(* IEC 61131-3 sources: sis-interlock-demo/src/GVLs/Generated, 3 files *)

(* ---- GVL_Sis.gvl.st ---- *)
// AUTO-GENERATED by cemgen 1.0.0 — не редактировать: правьте матрицу и запустите
//   python -m cemgen generate <файл матрицы .csv или .xlsx>
// Матрица: SIS-V101-CEM, объект V-101, ревизия B от 2026-10-19, SHA-256 сетки df2ed4841a9453ca
// Назначение: экземпляры ПАЗ объекта V-101: источник времени, журнал событий, приложение ПАЗ и
//             команды HMI (ST_SisCmd). Вызов — PRG_Sis.
// Автор:      kr0nsch; код — генератор cemgen
// Версия:     1.0.0
// Документ:   docs/DESIGN.md, раздел «10. Генератор cemgen»; docs/cause_effect_matrix.md
// ВНИМАНИЕ:   код демонстрационный и не предназначен для систем безопасности. Реальная ПАЗ требует
//             определения SIL, сертифицированных аппаратных и программных средств и валидации по
//             ГОСТ Р МЭК 61511.
{attribute 'qualified_only'}
VAR_GLOBAL
    fbTime : PL.FB_SystemTime;   // монотонное время LTIME (PL.I_TimeSource)
    fbLog  : FB_SisEventLog;     // журнал событий ПАЗ, кольцо GVL_Const.SIS_LOG_SIZE
    fbApp  : FB_SisApp;          // ПАЗ объекта: привязка, голосование, матрица, выходы
    stCmd  : ST_SisCmd;          // команды HMI: сброс, пусковые обходы, байпасы каналов
END_VAR

(* ---- GVL_SisCfg.gvl.st ---- *)
// AUTO-GENERATED by cemgen 1.0.0 — не редактировать: правьте матрицу и запустите
//   python -m cemgen generate <файл матрицы .csv или .xlsx>
// Матрица: SIS-V101-CEM, объект V-101, ревизия B от 2026-10-19, SHA-256 сетки df2ed4841a9453ca
// Назначение: конфигурация ПАЗ объекта V-101 из матрицы причин и следствий: номера причин и
//             следствий, шкалы датчиков, матрица CEM_CFG (с CRC) и группы голосования VOTE_CFG.
//             VAR_GLOBAL CONSTANT: с HMI не меняется (решение D-09), правка — только через матрицу
//             и генератор.
// Автор:      kr0nsch; код — генератор cemgen
// Версия:     1.0.0
// Документ:   docs/DESIGN.md, раздел «10. Генератор cemgen»; docs/cause_effect_matrix.md
// ВНИМАНИЕ:   код демонстрационный и не предназначен для систем безопасности. Реальная ПАЗ требует
//             определения SIL, сертифицированных аппаратных и программных средств и валидации по
//             ГОСТ Р МЭК 61511.
{attribute 'qualified_only'}
VAR_GLOBAL CONSTANT
    // Номера причин: индекс i строки матрицы, бит маски i − 1
    CAUSE_PSHH101       : UINT := 1;   // Давление в V-101 аварийно высокое
    CAUSE_PSLL101       : UINT := 2;   // Давление в V-101 аварийно низкое
    CAUSE_LSHH102       : UINT := 3;   // Уровень жидкости в V-101 аварийно высокий
    CAUSE_LSLL102       : UINT := 4;   // Уровень жидкости в V-101 аварийно низкий
    CAUSE_TSHH103       : UINT := 5;   // Температура жидкости в V-101 аварийно высокая
    CAUSE_ASHH104       : UINT := 6;   // Загазованность у V-101 аварийно высокая
    CAUSE_BSH105        : UINT := 7;   // Пожар у V-101
    CAUSE_HS106         : UINT := 8;   // Аварийный останов кнопкой
    CAUSE_PSLL108       : UINT := 9;   // Давление воздуха КИП аварийно низкое
    CAUSE_ESL109        : UINT := 10;   // Потеря напряжения щита 0,4 кВ
    CAUSE_COUNT         : UINT := 10;   // причин в матрице
    // Номера следствий: индекс j столбца матрицы
    EFFECT_ESDV101      : UINT := 1;   // Клапан-отсекатель на входе V-101
    EFFECT_BDV101       : UINT := 2;   // Клапан аварийного сброса давления на факел
    EFFECT_ESDV102      : UINT := 3;   // Клапан-отсекатель на линии нефти
    EFFECT_P101A        : UINT := 4;   // Насос откачки нефти P-101A
    EFFECT_P101B        : UINT := 5;   // Насос откачки нефти P-101B
    EFFECT_H101         : UINT := 6;   // Погружной электронагреватель H-101 в V-101
    EFFECT_UA110        : UINT := 7;   // Общая сигнализация «Срабатывание ПАЗ»
    EFFECT_COUNT        : UINT := 7;   // следствий в матрице
    // Шкалы датчиков 4–20 мА (инж. ед.) и нормальные токи для демо и тестов
    AI_PT101A_LO_EU     : REAL := 0.0;   // PT101A: шкала 0…1,6 МПа
    AI_PT101A_HI_EU     : REAL := 1.6;
    AI_PT101A_NORMAL_MA : REAL := 10.0;   // 0,6 МПа
    AI_PT101B_LO_EU     : REAL := 0.0;   // PT101B: шкала 0…1,6 МПа
    AI_PT101B_HI_EU     : REAL := 1.6;
    AI_PT101B_NORMAL_MA : REAL := 10.0;   // 0,6 МПа
    AI_PT101C_LO_EU     : REAL := 0.0;   // PT101C: шкала 0…1,6 МПа
    AI_PT101C_HI_EU     : REAL := 1.6;
    AI_PT101C_NORMAL_MA : REAL := 10.0;   // 0,6 МПа
    AI_LT102A_LO_EU     : REAL := 0.0;   // LT102A: шкала 0…2,4 м
    AI_LT102A_HI_EU     : REAL := 2.4;
    AI_LT102A_NORMAL_MA : REAL := 12.0;   // 1,2 м
    AI_LT102B_LO_EU     : REAL := 0.0;   // LT102B: шкала 0…2,4 м
    AI_LT102B_HI_EU     : REAL := 2.4;
    AI_LT102B_NORMAL_MA : REAL := 12.0;   // 1,2 м
    AI_LT102C_LO_EU     : REAL := 0.0;   // LT102C: шкала 0…2,4 м
    AI_LT102C_HI_EU     : REAL := 2.4;
    AI_LT102C_NORMAL_MA : REAL := 12.0;   // 1,2 м
    AI_TT103A_LO_EU     : REAL := 0.0;   // TT103A: шкала 0…150 °C
    AI_TT103A_HI_EU     : REAL := 150.0;
    AI_TT103A_NORMAL_MA : REAL := 10.4;   // 60 °C
    AI_TT103B_LO_EU     : REAL := 0.0;   // TT103B: шкала 0…150 °C
    AI_TT103B_HI_EU     : REAL := 150.0;
    AI_TT103B_NORMAL_MA : REAL := 10.4;   // 60 °C
    AI_AT104A_LO_EU     : REAL := 0.0;   // AT104A: шкала 0…100 % НКПР
    AI_AT104A_HI_EU     : REAL := 100.0;
    AI_AT104A_NORMAL_MA : REAL := 4.0;   // 0 % НКПР
    AI_AT104B_LO_EU     : REAL := 0.0;   // AT104B: шкала 0…100 % НКПР
    AI_AT104B_HI_EU     : REAL := 100.0;
    AI_AT104B_NORMAL_MA : REAL := 4.0;   // 0 % НКПР
    AI_AT104C_LO_EU     : REAL := 0.0;   // AT104C: шкала 0…100 % НКПР
    AI_AT104C_HI_EU     : REAL := 100.0;
    AI_AT104C_NORMAL_MA : REAL := 4.0;   // 0 % НКПР
    // Матрица причин и следствий (DESIGN.md, 4.2, 6.8): маска следствия — «X» в его столбце
    CEM_CFG : ST_CemCfg := (uiCauseCount := 10, uiEffectCount := 7, xStartTripped := TRUE,
        wMatrixCrc := 16#CD40,
        astCause := [
            (xEnable := TRUE, eSource := E_CauseSource.Voting, tDelay := T#2S),                 // 1 PSHH101
            (xEnable := TRUE, eSource := E_CauseSource.Voting, tDelay := T#5S,
                xOverrideAllowed := TRUE, tOverrideMax := T#15M, tOverrideClear := T#30S),      // 2 PSLL101
            (xEnable := TRUE, eSource := E_CauseSource.Voting, tDelay := T#3S),                 // 3 LSHH102
            (xEnable := TRUE, eSource := E_CauseSource.Voting, tDelay := T#5S,
                xOverrideAllowed := TRUE, tOverrideMax := T#30M, tOverrideClear := T#1M),       // 4 LSLL102
            (xEnable := TRUE, eSource := E_CauseSource.Voting, tDelay := T#5S),                 // 5 TSHH103
            (xEnable := TRUE, eSource := E_CauseSource.Voting, tDelay := T#2S),                 // 6 ASHH104
            (xEnable := TRUE, eSource := E_CauseSource.Voting, tDelay := T#0S),                 // 7 BSH105
            (xEnable := TRUE, eSource := E_CauseSource.Voting, tDelay := T#0S),                 // 8 HS106
            (xEnable := TRUE, eSource := E_CauseSource.Voting, tDelay := T#10S,
                xOverrideAllowed := TRUE, tOverrideMax := T#10M, tOverrideClear := T#30S),      // 9 PSLL108
            (xEnable := TRUE, eSource := E_CauseSource.Voting, tDelay := T#2S),                 // 10 ESL109
            (xEnable := FALSE),                                                                 // 11 — резерв
            (xEnable := FALSE),                                                                 // 12 — резерв
            (xEnable := FALSE),                                                                 // 13 — резерв
            (xEnable := FALSE),                                                                 // 14 — резерв
            (xEnable := FALSE),                                                                 // 15 — резерв
            (xEnable := FALSE)],                                                                // 16 — резерв
        astEffect := [
            (eSafeState := E_SafeState.Closed, wCauseMask := 16#01E7),         // 1 ESDV101: 1, 2, 3, 6, 7, 8, 9
            (eSafeState := E_SafeState.Open, wCauseMask := 16#00C0),           // 2 BDV101: 7, 8
            (eSafeState := E_SafeState.Closed, wCauseMask := 16#01EA),         // 3 ESDV102: 2, 4, 6, 7, 8, 9
            (eSafeState := E_SafeState.Stopped, wCauseMask := 16#03EA),        // 4 P101A: 2, 4, 6, 7, 8, 9, 10
            (eSafeState := E_SafeState.Stopped, wCauseMask := 16#03EA),        // 5 P101B: 2, 4, 6, 7, 8, 9, 10
            (eSafeState := E_SafeState.Off, wCauseMask := 16#03FF),            // 6 H101: 1, 2, 3, 4, 5, 6, 7, 8, 9, 10
            (eSafeState := E_SafeState.Alarm, wCauseMask := 16#03FF),          // 7 UA110: 1, 2, 3, 4, 5, 6, 7, 8, 9, 10
            (wCauseMask := 0),                                                 // 8 — резерв
            (wCauseMask := 0),                                                 // 9 — резерв
            (wCauseMask := 0),                                                 // 10 — резерв
            (wCauseMask := 0),                                                 // 11 — резерв
            (wCauseMask := 0),                                                 // 12 — резерв
            (wCauseMask := 0),                                                 // 13 — резерв
            (wCauseMask := 0),                                                 // 14 — резерв
            (wCauseMask := 0),                                                 // 15 — резерв
            (wCauseMask := 0)]);                                               // 16 — резерв
    // Группы голосования по причинам (DESIGN.md, 5); ext — без голосования (eArch := None)
    VOTE_CFG : ARRAY[1..GVL_Const.SIS_CAUSES_MAX] OF ST_VotingCfg := [
        (eArch := E_VoteArch.Vote2oo3, ePolicy := E_DegradePolicy.VoteTrip,
            eInput := E_SisInputKind.Analog, eLimitDir := E_LimitDir.High,
            rTripLimit_eu := 0.9, rHyst_eu := 0.02, rDiscrepancyMax_eu := 0.05,
            tDiscrepancyDelay := T#10S, tBypassMax := T#8H, uiMaxBypass := 1),                  // 1 PSHH101
        (eArch := E_VoteArch.Vote2oo3, ePolicy := E_DegradePolicy.VoteTrip,
            eInput := E_SisInputKind.Analog, eLimitDir := E_LimitDir.Low,
            rTripLimit_eu := 0.15, rHyst_eu := 0.02, rDiscrepancyMax_eu := 0.05,
            tDiscrepancyDelay := T#10S, tBypassMax := T#8H, uiMaxBypass := 1),                  // 2 PSLL101
        (eArch := E_VoteArch.Vote2oo3, ePolicy := E_DegradePolicy.DegradeAvailable,
            eInput := E_SisInputKind.Analog, eLimitDir := E_LimitDir.High,
            rTripLimit_eu := 1.8, rHyst_eu := 0.02, rDiscrepancyMax_eu := 0.1,
            tDiscrepancyDelay := T#10S, tBypassMax := T#8H, uiMaxBypass := 1),                  // 3 LSHH102
        (eArch := E_VoteArch.Vote2oo3, ePolicy := E_DegradePolicy.DegradeAvailable,
            eInput := E_SisInputKind.Analog, eLimitDir := E_LimitDir.Low,
            rTripLimit_eu := 0.5, rHyst_eu := 0.02, rDiscrepancyMax_eu := 0.1,
            tDiscrepancyDelay := T#10S, tBypassMax := T#8H, uiMaxBypass := 1),                  // 4 LSLL102
        (eArch := E_VoteArch.Vote1oo2, ePolicy := E_DegradePolicy.DegradeSafe,
            eInput := E_SisInputKind.Analog, eLimitDir := E_LimitDir.High,
            rTripLimit_eu := 85.0, rHyst_eu := 1.0, rDiscrepancyMax_eu := 5.0,
            tDiscrepancyDelay := T#10S, tBypassMax := T#8H, uiMaxBypass := 1),                  // 5 TSHH103
        (eArch := E_VoteArch.Vote2oo3, ePolicy := E_DegradePolicy.DegradeSafe,
            eInput := E_SisInputKind.Analog, eLimitDir := E_LimitDir.High,
            rTripLimit_eu := 50.0, rHyst_eu := 5.0, rDiscrepancyMax_eu := 10.0,
            tDiscrepancyDelay := T#30S, tBypassMax := T#8H, uiMaxBypass := 1),                  // 6 ASHH104
        (eArch := E_VoteArch.Vote1oo2, ePolicy := E_DegradePolicy.DegradeSafe,
            eInput := E_SisInputKind.Discrete, xDiHealthy := TRUE, tBypassMax := T#8H,
            uiMaxBypass := 1),                                                                  // 7 BSH105
        (eArch := E_VoteArch.Vote1oo2, ePolicy := E_DegradePolicy.VoteTrip,
            eInput := E_SisInputKind.Discrete, xDiHealthy := TRUE, tBypassMax := T#0S,
            uiMaxBypass := 0),                                                                  // 8 HS106
        (eArch := E_VoteArch.Vote2oo2, ePolicy := E_DegradePolicy.DegradeSafe,
            eInput := E_SisInputKind.Discrete, xDiHealthy := TRUE, tBypassMax := T#4H,
            uiMaxBypass := 1),                                                                  // 9 PSLL108
        (eArch := E_VoteArch.Vote1oo1, ePolicy := E_DegradePolicy.VoteTrip,
            eInput := E_SisInputKind.Discrete, xDiHealthy := TRUE, tBypassMax := T#0S,
            uiMaxBypass := 0),                                                                  // 10 ESL109
        (eArch := E_VoteArch.None),                                                             // 11 — резерв
        (eArch := E_VoteArch.None),                                                             // 12 — резерв
        (eArch := E_VoteArch.None),                                                             // 13 — резерв
        (eArch := E_VoteArch.None),                                                             // 14 — резерв
        (eArch := E_VoteArch.None),                                                             // 15 — резерв
        (eArch := E_VoteArch.None)];                                                            // 16 — резерв
END_VAR

(* ---- GVL_SisIo.gvl.st ---- *)
// AUTO-GENERATED by cemgen 1.0.0 — не редактировать: правьте матрицу и запустите
//   python -m cemgen generate <файл матрицы .csv или .xlsx>
// Матрица: SIS-V101-CEM, объект V-101, ревизия B от 2026-10-19, SHA-256 сетки df2ed4841a9453ca
// Назначение: образ ввода-вывода ПАЗ объекта V-101. Поля stIo привязываются к каналам модулей
//             ввода-вывода; в демо без ввода-вывода PRG_Main ставит нормальные значения
//             (F_SisIoNormal).
// Автор:      kr0nsch; код — генератор cemgen
// Версия:     1.0.0
// Документ:   docs/DESIGN.md, раздел «10. Генератор cemgen»; docs/cause_effect_matrix.md
// ВНИМАНИЕ:   код демонстрационный и не предназначен для систем безопасности. Реальная ПАЗ требует
//             определения SIL, сертифицированных аппаратных и программных средств и валидации по
//             ГОСТ Р МЭК 61511.
{attribute 'qualified_only'}
VAR_GLOBAL
    stIo : ST_SisIo;   // входы датчиков, ключи, кнопка, выходы-разрешения xQ*
END_VAR
